TYPE ST_PQ :		// P·Q 한 쌍 (유닛 지령·쓴 값·보정량 공통)
STRUCT
	fP			: REAL;		// kW, 방전·공급 +
	fQ			: REAL;		// kvar, 공급 +
END_STRUCT
END_TYPE

(* stored: Version 1.1.0.1, ProductVersion 3.1.4024.15
   DUT ST_PQ: Id {822e7d2c-0cbd-4444-834e-af13fefd24b4} *)
